Fanuc KAREL source: kt00710.KL

-- PROVISIONAL review KL for V940-1; original PC SHA256 181f7c32f5a8f55b6ba7338977758f61bae91e818d8a66ab36ee69ef1abc2910
-- Incomplete behavior may be omitted. Consult companion uncertainty JSON. Do not deploy.
PROGRAM KT00710
%NOLOCKGROUP
VAR
  B1 : BOOLEAN
  B2 : BOOLEAN
  OUT : BOOLEAN
BEGIN
  -- V9_ZERO_TABLE_METADATA_HINT layout=0001; no indexed target words; source/name/runtime held
  -- UNRESOLVED_PC offsets 5-12; opcodes 9D,23
  -- UNRESOLVED_PC offsets 17-24; opcodes 9C,23
  -- UNRESOLVED_PC offsets 29-36; opcodes 9D,23
  -- UNRESOLVED_PC offsets 41-48; opcodes 9C,23
  -- UNRESOLVED_PC offsets 53-68; opcodes 22,63,23
  -- UNRESOLVED_PC offsets 73-77; opcodes 7F
END KT00710
